(* Logix 5000 project; controller SmartManufacturingCell Emulate 5570 rev 33.11; software revision 33.03; part 5 of 5 *)
(* tags used below, declared in another part *)
   AutoRequestONS : BOOL;
   ConfigurationValid : BOOL;
   ManualRequestONS : BOOL;
   ModeChangeAllowed : BOOL;
   Recovery_CommandsReleased : BOOL;
   Recovery_PhaseClear : BOOL;
   Recovery_SensorsClear : BOOL;
   Recovery_TrackingClear : BOOL;
   Start_CommandsReleased : BOOL;
   Start_EquipmentReady : BOOL;
   StartRequestONS : BOOL;
   Startup_CheckPending : BOOL;
   Cfg_FillTimeMs : DINT;   // Fill duration; 100..3000 ms. Sampled when filling starts.
   Cfg_InspectionTimeMs : DINT;   // Inspection duration; 100..2000 ms. Sampled when inspection starts.
   Conveyor_Flt_FailToStart : BOOL;   // Conveyor commanded but running feedback missing for 2 s Latched; clear cell, remove cause, then fresh Reset.
   Conveyor_Sts_ResetAccepted : BOOL;   // One-execution indication that conveyor fault reset was accepted.
   Exit_Flt_DischargeTimeout : BOOL;   // Good or reject bottle departure not confirmed within 3 s Latched; clear cell, remove cause, then fresh Reset.
   Exit_Sts_ResetAccepted : BOOL;   // Exit Sts ResetAccepted
   Exit_Sts_State : DINT;   // 0 Empty; 10 Waiting; 20 Good discharge; 30 Extending; 40 Reject discharge; 50 Retracting; 60 Complete; 90 Faulted
   Filling_Flt_FillTimeout : BOOL;   // Fill completion not received within 4 s Latched; clear cell, remove cause, then fresh Reset.
   Filling_Flt_ValveFailToClose : BOOL;   // Fill valve did not close within 2 s Latched; clear cell, remove cause, then fresh Reset.
   Filling_Sts_ResetAccepted : BOOL;   // Filling Sts ResetAccepted
   Filling_Sts_State : DINT;   // 0 Empty; 10 Waiting; 20 Filling; 30 Closing; 40 Complete; 90 Faulted
   HMI_Cmd_ClearCell : BOOL;   // Request removal of simulated bottles during fault recovery
   HMI_Cmd_ConveyorJog : BOOL;   // Request conveyor movement while held
   HMI_Cmd_FillValveOpen : BOOL;
   HMI_Cmd_LoadBottle : BOOL;   // Request one simulated bottle at the available entry position
   HMI_Cmd_RejectExtend : BOOL;
   HMI_Cmd_Reset : BOOL;   // Request fault reset after recovery conditions are satisfied
   HMI_Cmd_SelectAuto : BOOL;   // Request Auto mode
   HMI_Cmd_SelectManual : BOOL;   // Request Manual mode
   HMI_Cmd_Start : BOOL;   // Request automatic production start
   HMI_Cmd_Stop : BOOL;   // Request controlled production stop
   HMI_Sim_BottleMissingAtFill : BOOL;   // Suppress Fill photoeye while retaining simulated bottle presence. Simulation test only.
   HMI_Sim_ConveyorFailToStart : BOOL;   // Suppress conveyor running feedback. Simulation test only.
   HMI_Sim_FillFailToComplete : BOOL;   // Suppress simulated filling completion. Simulation test only.
   HMI_Sim_FillValveFailToClose : BOOL;   // Suppress fill valve closed feedback. Simulation test only.
   HMI_Sim_GoodDischargeJam : BOOL;   // Prevent good bottle departure. Simulation test only.
   HMI_Sim_IndexJam : BOOL;   // Prevent simulated index travel from completing. Simulation test only.
   HMI_Sim_IndexPositionMismatch : BOOL;   // Invert simulated Fill occupancy on transfer to test confirmation. Simulation test only.
   HMI_Sim_InspectionFailToComplete : BOOL;   // Prevent inspection process timer from completing. Simulation test only.
   HMI_Sim_RejectDischargeJam : BOOL;   // Prevent rejected bottle departure. Simulation test only.
   HMI_Sim_RejectFailToExtend : BOOL;   // Suppress reject extended feedback. Simulation test only.
   HMI_Sim_RejectFailToRetract : BOOL;   // Suppress reject retracted feedback. Simulation test only.
   Inspection_Flt_Timeout : BOOL;   // Inspection did not finish within 3 s Latched; clear cell, remove cause, then fresh Reset.
   Inspection_Sts_ResetAccepted : BOOL;   // Inspection Sts ResetAccepted
   Inspection_Sts_State : DINT;   // 0 Empty; 10 Waiting; 20 Inspecting; 40 Complete; 90 Faulted
   Production_Bottles : UDT_Bottle[4];
   Production_Flt_IndexConfirmTimeout : BOOL;   // Post-index positions not confirmed within 1 s Latched; clear cell, remove cause, then fresh Reset.
   Production_Flt_IndexInterlock : BOOL;   // Movement interlock lost during indexing Latched; clear cell, remove cause, then fresh Reset.
   Production_Flt_IndexTimeout : BOOL;   // Index completion not received within 3 s Latched; clear cell, remove cause, then fresh Reset.
   Production_Flt_InvalidConfiguration : BOOL;   // Fill or inspection time outside permitted limits Latched; clear cell, remove cause, then fresh Reset.
   Production_Flt_InvalidState : BOOL;   // Machine, sequence, station state, or mode combination invalid Latched; clear cell, remove cause, then fresh Reset.
   Production_Flt_StartupRecoveryRequired : BOOL;   // Restart found bottles or interrupted activity Latched; clear cell, remove cause, then fresh Reset.
   Production_Flt_TrackingMismatch : BOOL;   // Stationary bottle tracking and sensors disagree or processing history invalid Latched; clear cell, remove cause, then fr
   Production_Sts_ResetAccepted : BOOL;
   Production_Sts_SequenceState : DINT;   // 0 = Idle 10 = ProcessStations 20 = Indexing 30 = ConfirmPositions
   Reject_Flt_FailToExtend : BOOL;   // Reject actuator did not extend within 2 s Latched; clear cell, remove cause, then fresh Reset.
   Reject_Flt_FailToRetract : BOOL;   // Reject actuator did not retract within 2 s Latched; clear cell, remove cause, then fresh Reset.
   Reject_Sts_ResetAccepted : BOOL;
   Sim_In_ConveyorRunning : BOOL;   // Simulated conveyor movement feedback
   Sim_In_EntryPE : BOOL;   // Simulated bottle detected at entry
   Sim_In_ExitPE : BOOL;   // Simulated bottle detected at Reject/Exit position
   Sim_In_FillPE : BOOL;   // Simulated bottle detected at filling position
   Sim_In_FillValveClosed : BOOL;   // Simulated fill valve confirmed closed
   Sim_In_GoodExitPE : BOOL;   // Bottle detected passing through good discharge path
   Sim_In_IndexComplete : BOOL;   // Simulated conveyor completed one station-spacing movement
   Sim_In_InspectionPE : BOOL;   // Simulated bottle detected at inspection position
   Sim_In_RejectExitPE : BOOL;   // Bottle detected passing through reject discharge path
   Sim_In_RejectExtended : BOOL;   // Simulated reject actuator confirmed extended
   Sim_In_RejectRetracted : BOOL;   // Simulated reject actuator confirmed retracted
   Sim_Out_ConveyorRun : BOOL;   // Command simulated conveyor to run
   Sim_Out_FillValveOpen : BOOL;   // Command simulated fill valve to open
   Sim_Out_GoodDischargeRun : BOOL;   // Command simulated good-bottle discharge mechanism to run
   Sim_Out_RejectExtend : BOOL;   // Command simulated reject actuator to extend
   Sim_Sts_BottlesPresent : BOOL;   // Sim Sts BottlesPresent
   Sys_Sts_AutoMode : BOOL;   // Auto mode accepted and active
   Sys_Sts_BlockingFault : BOOL;   // Active blocking fault prevents production and manual equipment operation.
   Sys_Sts_CellEmpty : BOOL;   // Sys Sts CellEmpty
   Sys_Sts_EquipmentHome : BOOL;   // Sys Sts EquipmentHome
   Sys_Sts_InjectionsClear : BOOL;   // Sys Sts InjectionsClear
   Sys_Sts_MachineState : DINT;   // 0 = Stopped 10 = Running 20 = Stopping 30 = Faulted
   Sys_Sts_ManualMode : BOOL;   // Manual mode accepted and active
   Sys_Sts_OperationsIdle : BOOL;   // Sys Sts OperationsIdle
   Sys_Sts_ResetAllowed : BOOL;   // Sys Sts ResetAllowed
   Sys_Sts_StartAllowed : BOOL;
   Sys_Sts_StartupReady : BOOL;   // Sys Sts StartupReady
(* Program_System, continued *)

ROUTINE Configuration_Control   (* ladder *)
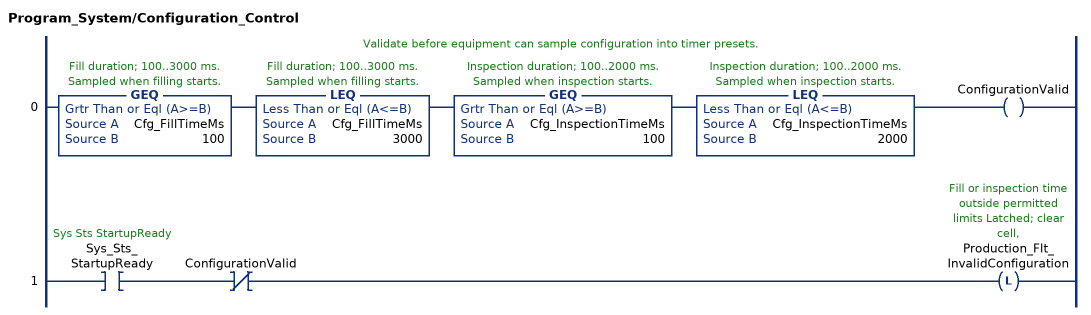
   // Validate before equipment can sample configuration into timer presets.
   0: GEQ(Cfg_FillTimeMs,100)LEQ(Cfg_FillTimeMs,3000)GEQ(Cfg_InspectionTimeMs,100)LEQ(Cfg_InspectionTimeMs,2000)OTE(ConfigurationValid);
   1: XIC(Sys_Sts_StartupReady)XIO(ConfigurationValid)OTL(Production_Flt_InvalidConfiguration);
END_ROUTINE

ROUTINE Fault_Control   (* ladder *)
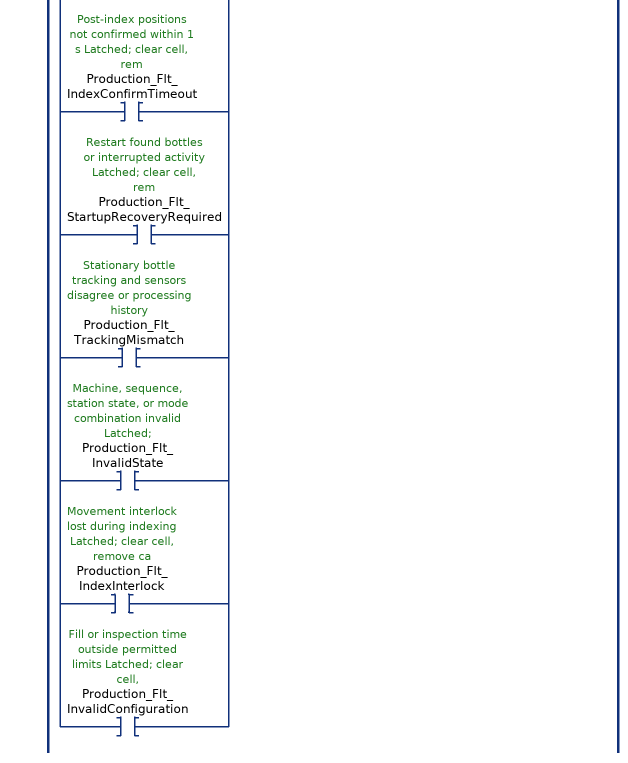
   0: [XIC(Conveyor_Flt_FailToStart) ,XIC(Filling_Flt_ValveFailToClose) ,XIC(Filling_Flt_FillTimeout) ,XIC(Inspection_Flt_Timeout) ,XIC(Reject_Flt_FailToExtend) ,XIC(Reject_Flt_FailToRetract) ,XIC(Exit_Flt_DischargeTimeout) ,XIC(Production_Flt_IndexTimeout) ,XIC(Production_Flt_IndexConfirmTimeout) ,XIC(Production_Flt_StartupRecoveryRequired) ,XIC(Production_Flt_TrackingMismatch) ,XIC(Production_Flt_InvalidState) ,XIC(Production_Flt_IndexInterlock) ,XIC(Production_Flt_InvalidConfiguration) ]OTE(Sys_Sts_BlockingFault);
END_ROUTINE

ROUTINE Machine_State   (* ladder *)
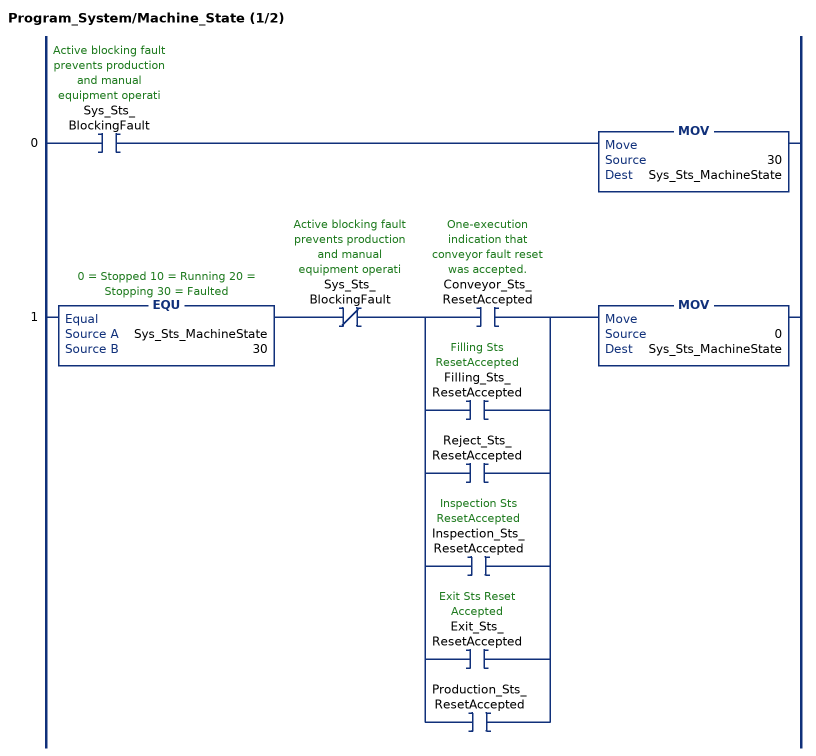
   0: XIC(Sys_Sts_BlockingFault)MOV(30,Sys_Sts_MachineState);
   1: EQU(Sys_Sts_MachineState,30)XIO(Sys_Sts_BlockingFault)[XIC(Conveyor_Sts_ResetAccepted) ,XIC(Filling_Sts_ResetAccepted) ,XIC(Reject_Sts_ResetAccepted) ,XIC(Inspection_Sts_ResetAccepted) ,XIC(Exit_Sts_ResetAccepted) ,XIC(Production_Sts_ResetAccepted) ]MOV(0,Sys_Sts_MachineState);
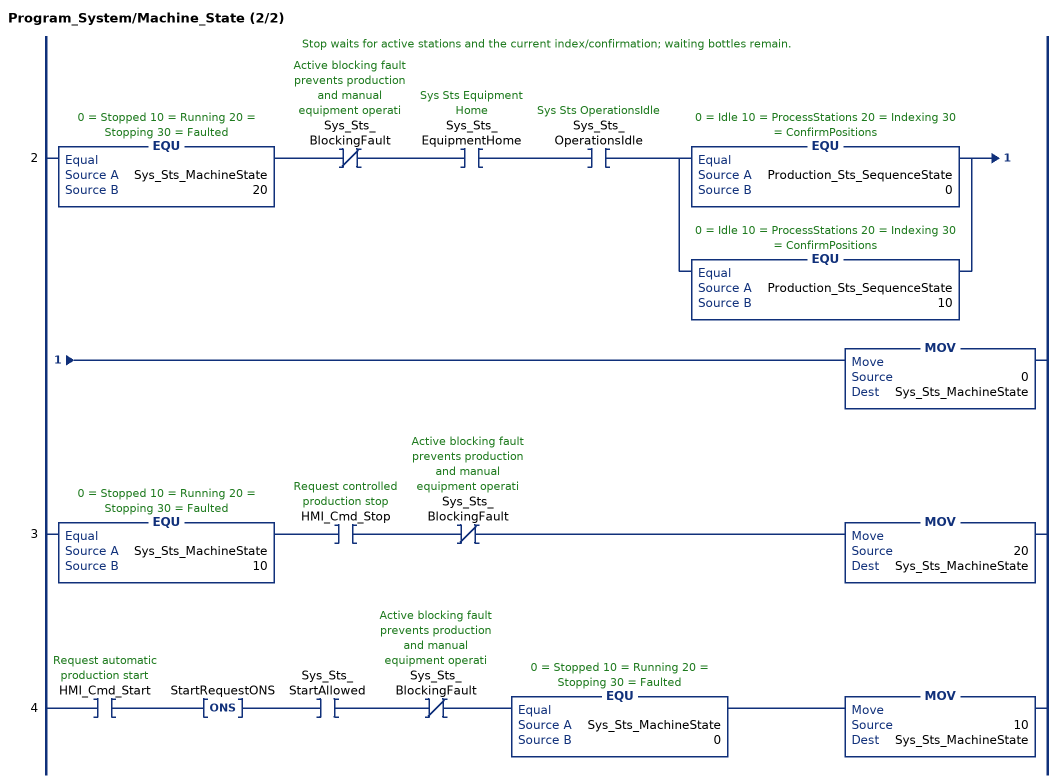
   // Stop waits for active stations and the current index/confirmation; waiting bottles remain.
   2: EQU(Sys_Sts_MachineState,20)XIO(Sys_Sts_BlockingFault)XIC(Sys_Sts_EquipmentHome)XIC(Sys_Sts_OperationsIdle)[EQU(Production_Sts_SequenceState,0) ,EQU(Production_Sts_SequenceState,10) ]MOV(0,Sys_Sts_MachineState);
   3: EQU(Sys_Sts_MachineState,10)XIC(HMI_Cmd_Stop)XIO(Sys_Sts_BlockingFault)MOV(20,Sys_Sts_MachineState);
   4: XIC(HMI_Cmd_Start)ONS(StartRequestONS)XIC(Sys_Sts_StartAllowed)XIO(Sys_Sts_BlockingFault)EQU(Sys_Sts_MachineState,0)MOV(10,Sys_Sts_MachineState);
END_ROUTINE

ROUTINE MainRoutine   (* ladder *)
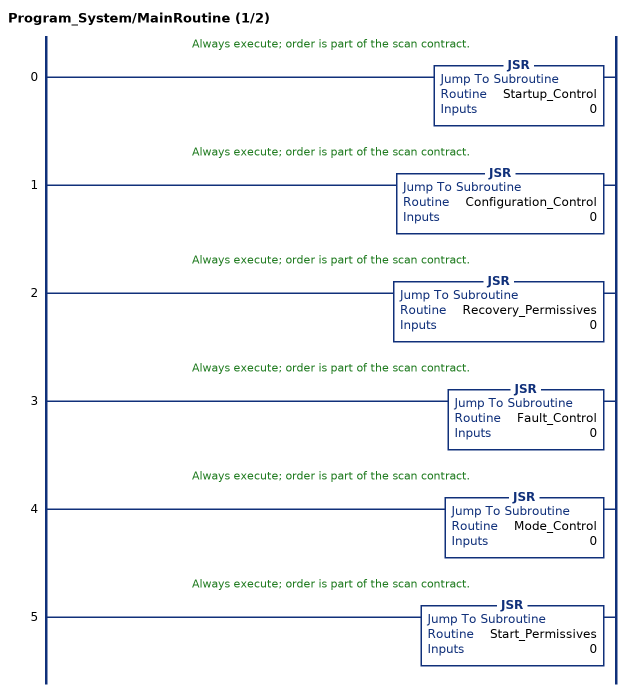
   // Always execute; order is part of the scan contract.
   0: JSR(Startup_Control,0);
   // Always execute; order is part of the scan contract.
   1: JSR(Configuration_Control,0);
   // Always execute; order is part of the scan contract.
   2: JSR(Recovery_Permissives,0);
   // Always execute; order is part of the scan contract.
   3: JSR(Fault_Control,0);
   // Always execute; order is part of the scan contract.
   4: JSR(Mode_Control,0);
   // Always execute; order is part of the scan contract.
   5: JSR(Start_Permissives,0);
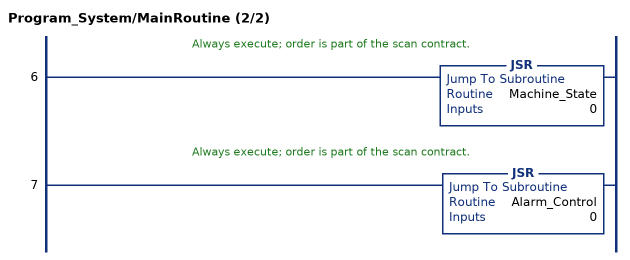
   // Always execute; order is part of the scan contract.
   6: JSR(Machine_State,0);
   // Always execute; order is part of the scan contract.
   7: JSR(Alarm_Control,0);
END_ROUTINE

ROUTINE Mode_Control   (* ladder *)
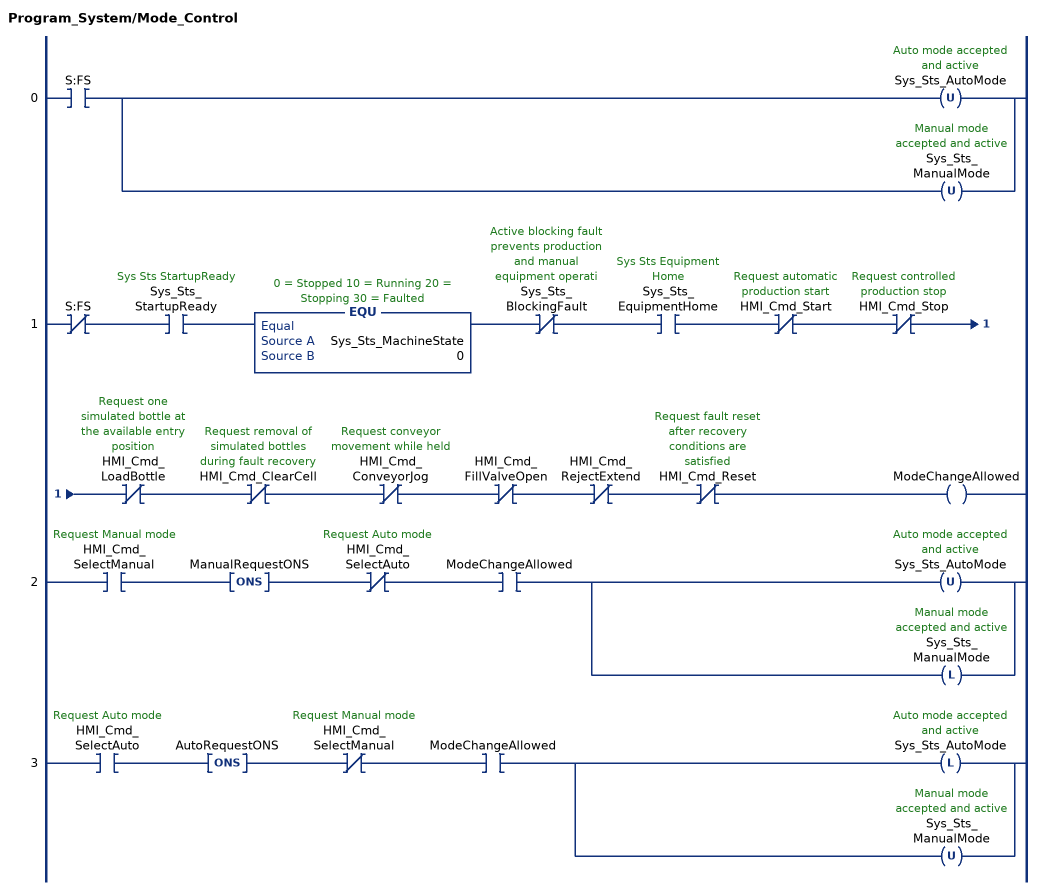
   0: XIC(S:FS)[OTU(Sys_Sts_AutoMode) ,OTU(Sys_Sts_ManualMode) ];
   1: XIO(S:FS)XIC(Sys_Sts_StartupReady)EQU(Sys_Sts_MachineState,0)XIO(Sys_Sts_BlockingFault)XIC(Sys_Sts_EquipmentHome)XIO(HMI_Cmd_Start)XIO(HMI_Cmd_Stop)XIO(HMI_Cmd_LoadBottle)XIO(HMI_Cmd_ClearCell)XIO(HMI_Cmd_ConveyorJog)XIO(HMI_Cmd_FillValveOpen)XIO(HMI_Cmd_RejectExtend)XIO(HMI_Cmd_Reset)OTE(ModeChangeAllowed);
   2: XIC(HMI_Cmd_SelectManual)ONS(ManualRequestONS)XIO(HMI_Cmd_SelectAuto)XIC(ModeChangeAllowed)[OTU(Sys_Sts_AutoMode) ,OTL(Sys_Sts_ManualMode) ];
   3: XIC(HMI_Cmd_SelectAuto)ONS(AutoRequestONS)XIO(HMI_Cmd_SelectManual)XIC(ModeChangeAllowed)[OTL(Sys_Sts_AutoMode) ,OTU(Sys_Sts_ManualMode) ];
END_ROUTINE

ROUTINE Recovery_Permissives   (* ladder *)
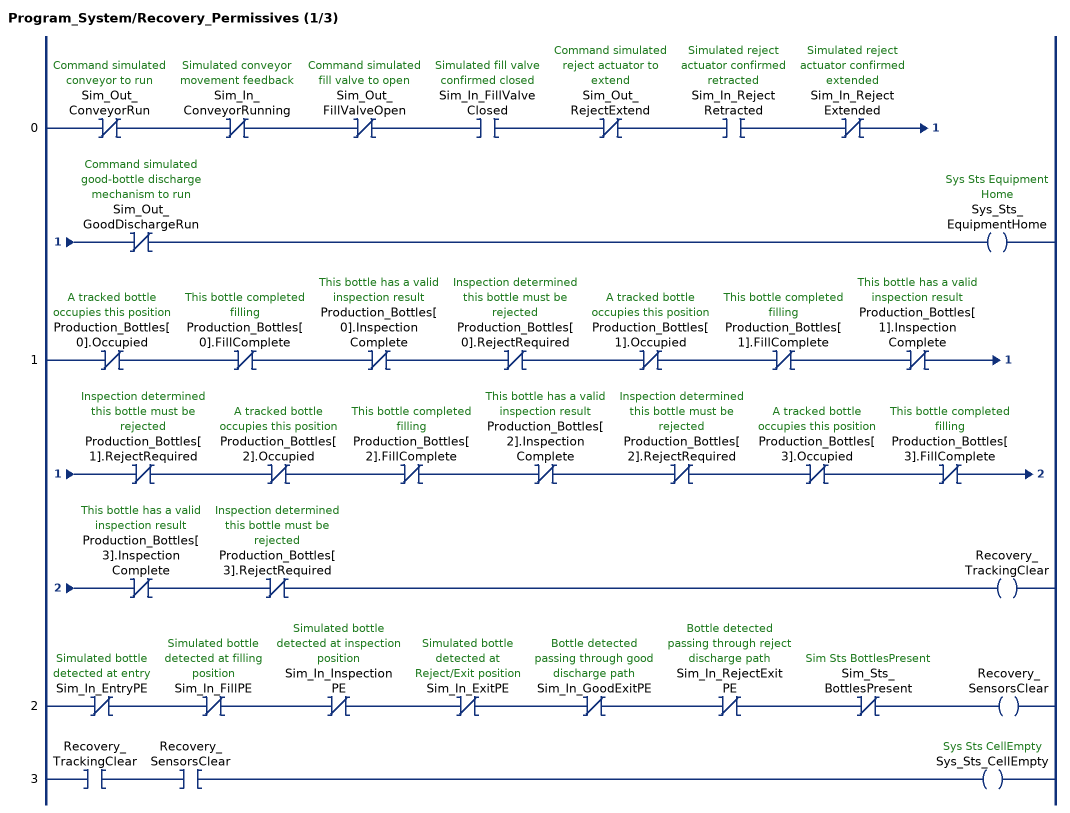
   0: XIO(Sim_Out_ConveyorRun)XIO(Sim_In_ConveyorRunning)XIO(Sim_Out_FillValveOpen)XIC(Sim_In_FillValveClosed)XIO(Sim_Out_RejectExtend)XIC(Sim_In_RejectRetracted)XIO(Sim_In_RejectExtended)XIO(Sim_Out_GoodDischargeRun)OTE(Sys_Sts_EquipmentHome);
   1: XIO(Production_Bottles[0].Occupied)XIO(Production_Bottles[0].FillComplete)XIO(Production_Bottles[0].InspectionComplete)XIO(Production_Bottles[0].RejectRequired)XIO(Production_Bottles[1].Occupied)XIO(Production_Bottles[1].FillComplete)XIO(Production_Bottles[1].InspectionComplete)XIO(Production_Bottles[1].RejectRequired)XIO(Production_Bottles[2].Occupied)XIO(Production_Bottles[2].FillComplete)XIO(Production_Bottles[2].InspectionComplete)XIO(Production_Bottles[2].RejectRequired)XIO(Production_Bottles[3].Occupied)XIO(Production_Bottles[3].FillComplete)XIO(Production_Bottles[3].InspectionComplete)XIO(Production_Bottles[3].RejectRequired)OTE(Recovery_TrackingClear);
   2: XIO(Sim_In_EntryPE)XIO(Sim_In_FillPE)XIO(Sim_In_InspectionPE)XIO(Sim_In_ExitPE)XIO(Sim_In_GoodExitPE)XIO(Sim_In_RejectExitPE)XIO(Sim_Sts_BottlesPresent)OTE(Recovery_SensorsClear);
   3: XIC(Recovery_TrackingClear)XIC(Recovery_SensorsClear)OTE(Sys_Sts_CellEmpty);
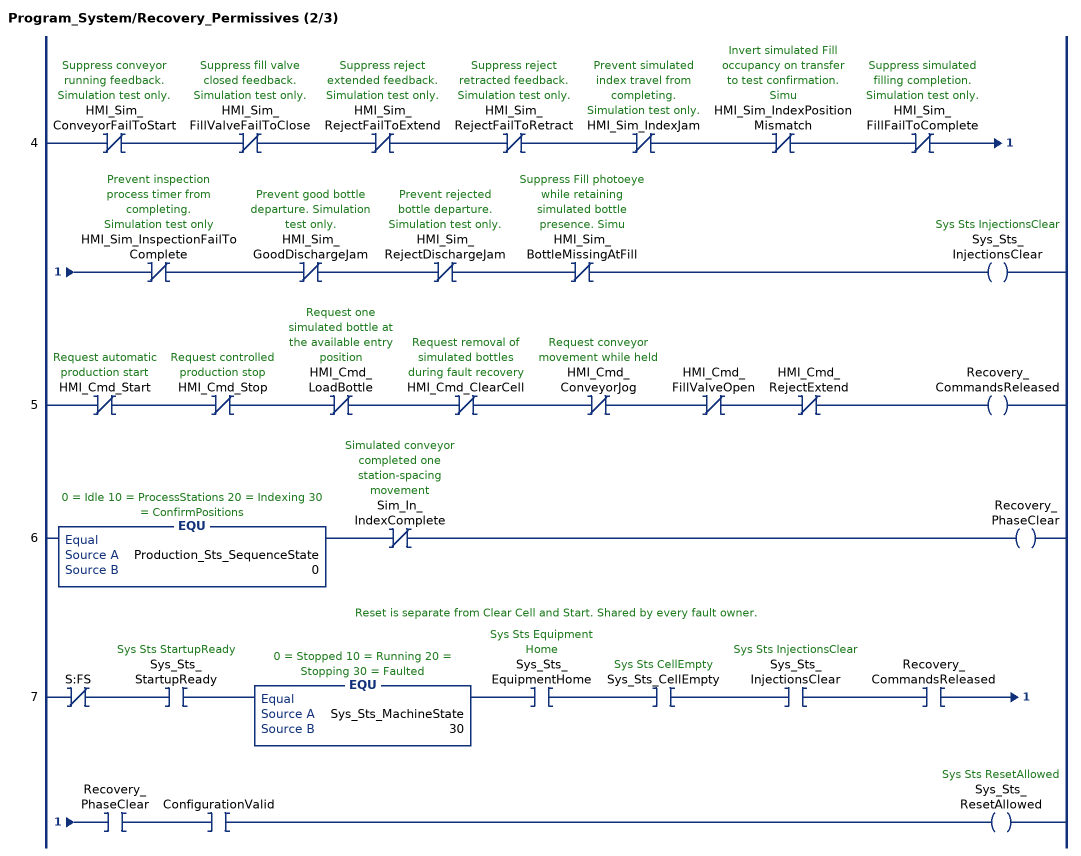
   4: XIO(HMI_Sim_ConveyorFailToStart)XIO(HMI_Sim_FillValveFailToClose)XIO(HMI_Sim_RejectFailToExtend)XIO(HMI_Sim_RejectFailToRetract)XIO(HMI_Sim_IndexJam)XIO(HMI_Sim_IndexPositionMismatch)XIO(HMI_Sim_FillFailToComplete)XIO(HMI_Sim_InspectionFailToComplete)XIO(HMI_Sim_GoodDischargeJam)XIO(HMI_Sim_RejectDischargeJam)XIO(HMI_Sim_BottleMissingAtFill)OTE(Sys_Sts_InjectionsClear);
   5: XIO(HMI_Cmd_Start)XIO(HMI_Cmd_Stop)XIO(HMI_Cmd_LoadBottle)XIO(HMI_Cmd_ClearCell)XIO(HMI_Cmd_ConveyorJog)XIO(HMI_Cmd_FillValveOpen)XIO(HMI_Cmd_RejectExtend)OTE(Recovery_CommandsReleased);
   6: EQU(Production_Sts_SequenceState,0)XIO(Sim_In_IndexComplete)OTE(Recovery_PhaseClear);
   // Reset is separate from Clear Cell and Start. Shared by every fault owner.
   7: XIO(S:FS)XIC(Sys_Sts_StartupReady)EQU(Sys_Sts_MachineState,30)XIC(Sys_Sts_EquipmentHome)XIC(Sys_Sts_CellEmpty)XIC(Sys_Sts_InjectionsClear)XIC(Recovery_CommandsReleased)XIC(Recovery_PhaseClear)XIC(ConfigurationValid)OTE(Sys_Sts_ResetAllowed);
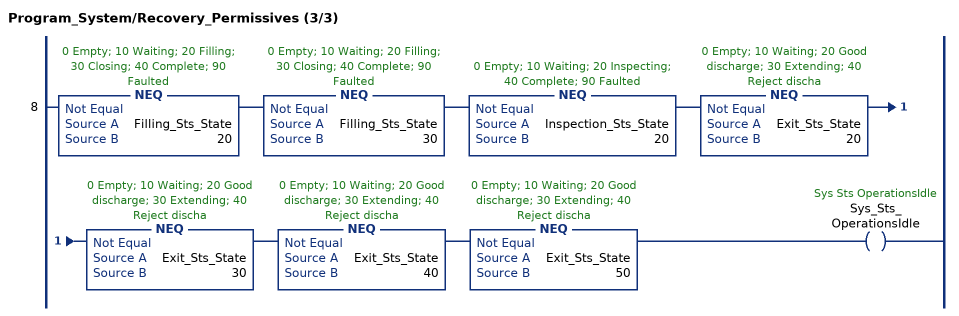
   8: NEQ(Filling_Sts_State,20)NEQ(Filling_Sts_State,30)NEQ(Inspection_Sts_State,20)NEQ(Exit_Sts_State,20)NEQ(Exit_Sts_State,30)NEQ(Exit_Sts_State,40)NEQ(Exit_Sts_State,50)OTE(Sys_Sts_OperationsIdle);
END_ROUTINE

ROUTINE Start_Permissives   (* ladder *)
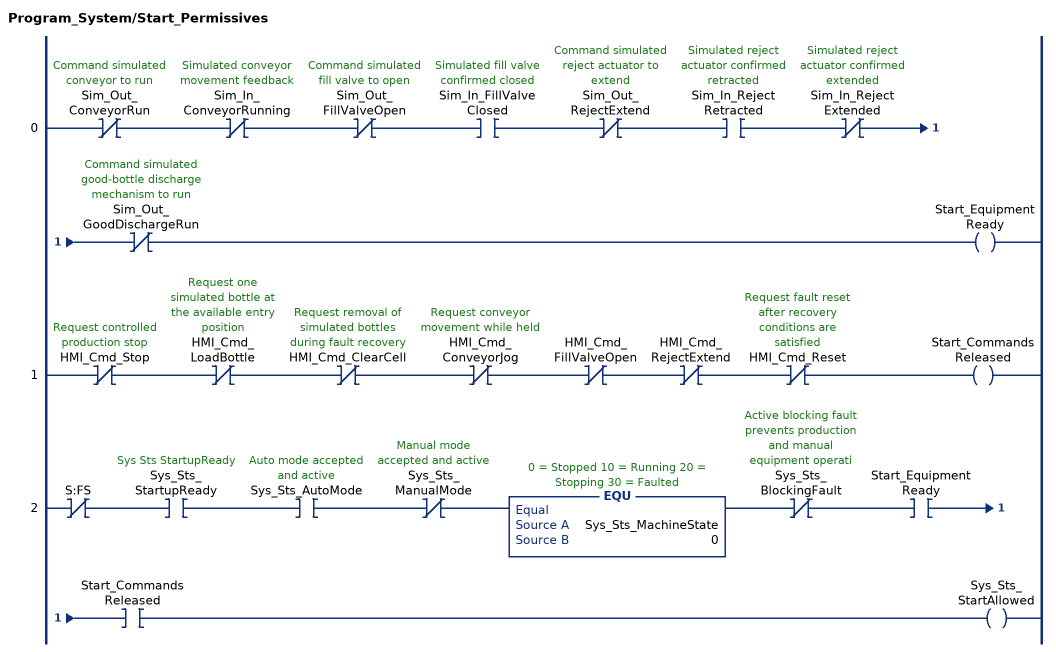
   0: XIO(Sim_Out_ConveyorRun)XIO(Sim_In_ConveyorRunning)XIO(Sim_Out_FillValveOpen)XIC(Sim_In_FillValveClosed)XIO(Sim_Out_RejectExtend)XIC(Sim_In_RejectRetracted)XIO(Sim_In_RejectExtended)XIO(Sim_Out_GoodDischargeRun)OTE(Start_EquipmentReady);
   1: XIO(HMI_Cmd_Stop)XIO(HMI_Cmd_LoadBottle)XIO(HMI_Cmd_ClearCell)XIO(HMI_Cmd_ConveyorJog)XIO(HMI_Cmd_FillValveOpen)XIO(HMI_Cmd_RejectExtend)XIO(HMI_Cmd_Reset)OTE(Start_CommandsReleased);
   2: XIO(S:FS)XIC(Sys_Sts_StartupReady)XIC(Sys_Sts_AutoMode)XIO(Sys_Sts_ManualMode)EQU(Sys_Sts_MachineState,0)XIO(Sys_Sts_BlockingFault)XIC(Start_EquipmentReady)XIC(Start_CommandsReleased)OTE(Sys_Sts_StartAllowed);
END_ROUTINE

ROUTINE Startup_Control   (* ladder *)
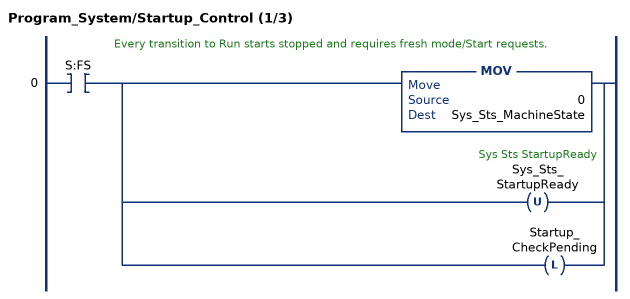
   // Every transition to Run starts stopped and requires fresh mode/Start requests.
   0: XIC(S:FS)[MOV(0,Sys_Sts_MachineState) ,OTU(Sys_Sts_StartupReady) ,OTL(Startup_CheckPending) ];
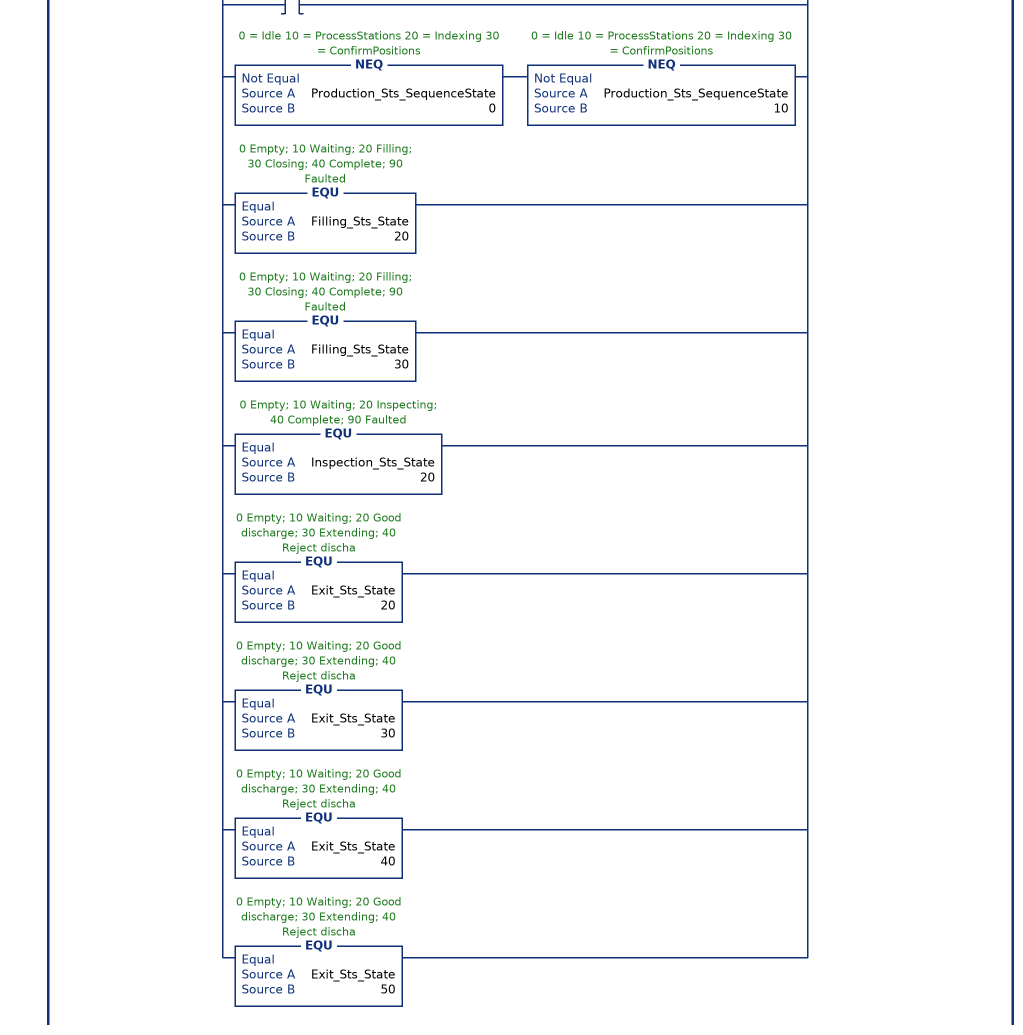
   // Wait one complete simulation pass: photoeyes are cleared by prescan. Physical presence also catches a masked sensor.
   1: XIC(Startup_CheckPending)XIO(S:FS)[XIC(Production_Bottles[0].Occupied) ,XIC(Production_Bottles[1].Occupied) ,XIC(Production_Bottles[2].Occupied) ,XIC(Production_Bottles[3].Occupied) ,XIC(Sim_In_EntryPE) ,XIC(Sim_In_FillPE) ,XIC(Sim_In_InspectionPE) ,XIC(Sim_In_ExitPE) ,XIC(Sim_In_GoodExitPE) ,XIC(Sim_In_RejectExitPE) ,XIC(Sim_Sts_BottlesPresent) ,NEQ(Production_Sts_SequenceState,0) NEQ(Production_Sts_SequenceState,10) ,[EQU(Filling_Sts_State,20) ,EQU(Filling_Sts_State,30) ] ,EQU(Inspection_Sts_State,20) ,[EQU(Exit_Sts_State,20) ,EQU(Exit_Sts_State,30) ,EQU(Exit_Sts_State,40) ,EQU(Exit_Sts_State,50) ] ]OTL(Production_Flt_StartupRecoveryRequired);
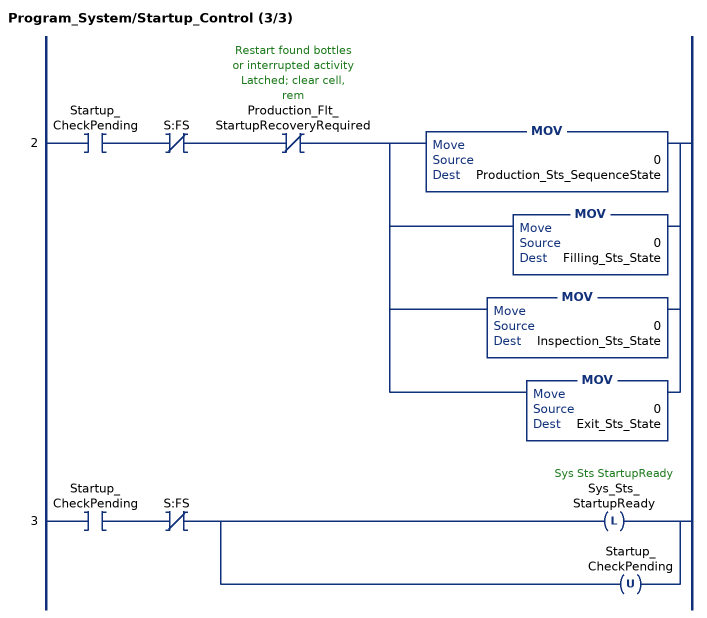
   2: XIC(Startup_CheckPending)XIO(S:FS)XIO(Production_Flt_StartupRecoveryRequired)[MOV(0,Production_Sts_SequenceState) ,MOV(0,Filling_Sts_State) ,MOV(0,Inspection_Sts_State) ,MOV(0,Exit_Sts_State) ];
   3: XIC(Startup_CheckPending)XIO(S:FS)[OTL(Sys_Sts_StartupReady) ,OTU(Startup_CheckPending) ];
END_ROUTINE
END_PROGRAM
